PROGRAM MAIN
VAR
    fbEnc : FB_SimEncoder;
    bGo   : BOOL;  // Wire to a HMI button or PLC tag
END_VAR

fbEnc(
    bActivate := bGo,
    rSpeed    := 1000.0,   // 1000 counts/s
    bDirection:= TRUE,
    nResolution := 4096    // e.g. 4096 PPR encoder
);

END_PROGRAM

(* stored: Version 1.1.0.1
   POU MAIN: Id {eb436a36-c8e2-4fab-9b6a-b8a59b9af6d9}, SpecialFunc None *)
